(*
	Owns the ended spans of every tracer created from it and hands them to processors.
	Stage the processors every scan, then call tick once; tick passes each ended span to
	every staged processor, releases the span, and clears the staged list.
	The sampler decides which ended spans reach the processors; see onEnd.

	Example:
	provider.stageProcessor(consoleProcessor);
	// ... tracers start and end spans ...
	provider.tick(failureReason => reason);
*)
FUNCTION_BLOCK FB_TracerProvider
VAR
	_resource: REFERENCE TO FB_Resource;  // borrowed; the declaring scope owns its lifetime
	_idGenerator: REFERENCE TO FB_IdGenerator_Base;  // borrowed; the declaring scope owns its lifetime
	_sampler: REFERENCE TO FB_Sampler;  // borrowed; the declaring scope owns its lifetime
	_spans: FB_SpanQueue(TcOtlp_GVL.MAX_SPAN_RECORDS_PER_SCAN);  // ended spans waiting to be processed
	_head: POINTER TO ST_LinkedListNode;  // staged processors; the nodes are owned, the processors borrowed
	_failureReason: E_TracerProviderFailureReason;  // first staging failure since the last tick
END_VAR
VAR_OUTPUT
	stagedProcessorCount: UDINT;
END_VAR

(* Releases the staged-list nodes. The processors themselves are borrowed and untouched. *)
METHOD _freeProcessors
VAR
	_idx: UDINT;
	_node: POINTER TO ST_LinkedListNode;
END_VAR
FOR _idx := 0 TO TcOtlp_GVL.MAX_LOOP_COUNT DO
	IF THIS^._head = 0 THEN
		EXIT;
	END_IF
	_node := THIS^._head^.nxt;
	__DELETE(THIS^._head);
	THIS^._head := _node;
	// count down per node, so the count never claims nodes that are gone or hides ones that remain
	IF THIS^.stagedProcessorCount > 0 THEN
		THIS^.stagedProcessorCount := THIS^.stagedProcessorCount - 1;
	END_IF
END_FOR
END_METHOD

METHOD FB_Exit : BOOL
VAR_INPUT
	bInCopyCode: BOOL;  // TRUE: the exit method is called in order to leave the instance which will be copied afterwards (online change).
END_VAR
IF NOT bInCopyCode THEN
	THIS^._freeProcessors();
END_IF
END_METHOD

//FB_Init is always available implicitly and it is used primarily for initialization.
//The return value is not evaluated. For a specific influence, you can also declare the
//methods explicitly and provide additional code there with the standard initialization
//code. You can evaluate the return value.
METHOD FB_Init: BOOL
VAR_INPUT
    bInitRetains: BOOL; // TRUE: the retain variables are initialized (reset warm / reset cold)
    bInCopyCode: BOOL;  // TRUE: the instance will be copied to the copy code afterward (online change)
	resource: REFERENCE TO FB_Resource;
	idGenerator: REFERENCE TO FB_IdGenerator_Base;  // the source of identifiers for every tracer of this provider
	sampler: REFERENCE TO FB_Sampler;  // decides which spans are sampled; TcOtlp_GVL.defaultSampler is the OpenTelemetry default
END_VAR
THIS^._resource REF= resource;
THIS^._idGenerator REF= idGenerator;
THIS^._sampler REF= sampler;
END_METHOD

(*
	Takes ownership of an ended span and queues it for processing. On success pSpan is
	cleared; on failure it is left unchanged and still owned by the caller.
	A span that is not sampled is released instead, and that counts as success. The sampler's
	onEnd is asked only about spans that are still sampled, so it can drop a span but never
	keep one that its onStart dropped.
*)
METHOD onEnd : BOOL
VAR_IN_OUT
	pSpan: POINTER TO FB_Span;
END_VAR
VAR
	_pushFailureReason: E_SpanQueueFailureReason;
END_VAR
IF pSpan = 0 THEN
	RETURN;
END_IF

IF pSpan^.isSampled() THEN
	THIS^.sampler.onEnd(span:=pSpan^);
END_IF

IF NOT pSpan^.isSampled() THEN
	pSpan^.delete(pSelf:=pSpan);
	onEnd := TRUE;
	RETURN;
END_IF

onEnd := THIS^._spans.push(pValue:=pSpan, failureReason=>_pushFailureReason);
END_METHOD

(*
	Adds a processor for the next tick. The processor is borrowed and must outlive the tick.
	Staging the same processor twice has no effect. At most MAX_LOOP_COUNT processors can be
	staged per tick; staging more fails with STAGE_PROCESSOR_FAILURE. Returns the provider so
	calls can chain.
*)
METHOD stageProcessor : REFERENCE TO FB_TracerProvider
VAR_INPUT
	processor: REFERENCE TO FB_SpanProcessor_Base;
END_VAR
VAR
	_idx: UDINT;
	_node: POINTER TO ST_LinkedListNode;
END_VAR
stageProcessor REF= THIS^;

IF NOT __ISVALIDREF(processor) THEN
	RETURN;
END_IF

IF THIS^._head = 0 THEN
	THIS^._head := __NEW(ST_LinkedListNode);
	IF THIS^._head = 0 THEN
		THIS^._failureReason := E_TracerProviderFailureReason.STAGE_PROCESSOR_FAILURE;
		RETURN;
	END_IF
	THIS^._head^.val := processor.pSelf;
	THIS^.stagedProcessorCount := 1;
	RETURN;
END_IF

_node := THIS^._head;
FOR _idx := 0 TO TcOtlp_GVL.MAX_LOOP_COUNT DO
	IF _node^.val = processor.pSelf THEN
		RETURN;
	ELSIF _node^.nxt = 0 THEN
		// at most MAX_LOOP_COUNT nodes, so _freeProcessors always releases them all
		IF THIS^.stagedProcessorCount >= TcOtlp_GVL.MAX_LOOP_COUNT THEN
			THIS^._failureReason := E_TracerProviderFailureReason.STAGE_PROCESSOR_FAILURE;
			RETURN;
		END_IF
		_node^.nxt := __NEW(ST_LinkedListNode);
		IF _node^.nxt = 0 THEN
			THIS^._failureReason := E_TracerProviderFailureReason.STAGE_PROCESSOR_FAILURE;
			RETURN;
		END_IF
		_node^.nxt^.val := processor.pSelf;
		THIS^.stagedProcessorCount := THIS^.stagedProcessorCount + 1;
		RETURN;
	END_IF
	_node := _node^.nxt;
END_FOR
END_METHOD

(*
	Call once per scan, after staging processors. Passes every queued ended span to each staged
	processor in staging order, releases the span, then ticks the processors and the id
	generator. The queue and the staged list are always cleared, so spans are never carried
	into the next scan: with no processors staged they are released unprocessed.
*)
METHOD tick : BOOL
VAR_OUTPUT
	failureReason: E_TracerProviderFailureReason;
END_VAR
VAR
	_i: UDINT;
	_j: UDINT;
	_count: UDINT;
	_node: POINTER TO ST_LinkedListNode;
	_processor: POINTER TO FB_SpanProcessor_Base;
	_span: POINTER TO FB_Span;
	_popFailureReason: E_SpanQueueFailureReason;
	_idGenFailureReason: E_IdGenFailureReason;
END_VAR
failureReason := THIS^._failureReason;
IF failureReason <> E_TracerProviderFailureReason.NA THEN
	JMP _endLabel;
END_IF

// hand each ended span to every staged processor, then release it
_count := THIS^._spans.count;
FOR _i := 1 TO _count DO
	IF NOT THIS^._spans.pop(pValue:=_span, failureReason=>_popFailureReason) THEN
		failureReason := E_TracerProviderFailureReason.QUEUE_POP_FAILURE;
		JMP _endLabel;
	END_IF
	_node := THIS^._head;
	FOR _j := 1 TO THIS^.stagedProcessorCount DO
		IF _node = 0 THEN
			failureReason := E_TracerProviderFailureReason.UNEXPECTED_NULL_LINKED_LIST_NODE;
			JMP _endLabel;
		END_IF
		_processor := _node^.val;
		IF _processor = 0 THEN
			failureReason := E_TracerProviderFailureReason.UNEXPECTED_NULL_PROCESSOR_POINTER;
			JMP _endLabel;
		END_IF
		_processor^.onEnd(_span^);
		_node := _node^.nxt;
	END_FOR
	_span^.delete(pSelf:=_span);
END_FOR

// tick each processor
_node := THIS^._head;
FOR _j := 1 TO THIS^.stagedProcessorCount DO
	IF _node = 0 THEN
		failureReason := E_TracerProviderFailureReason.UNEXPECTED_NULL_LINKED_LIST_NODE;
		JMP _endLabel;
	END_IF
	_processor := _node^.val;
	IF _processor = 0 THEN
		failureReason := E_TracerProviderFailureReason.UNEXPECTED_NULL_PROCESSOR_POINTER;
		JMP _endLabel;
	END_IF
	_processor^.tick();
	_node := _node^.nxt;
END_FOR

_endLabel:
IF _span <> 0 THEN _span^.delete(pSelf:=_span); END_IF
THIS^._spans.free();
THIS^._freeProcessors();
THIS^._failureReason := E_TracerProviderFailureReason.NA;

// refill the identifier buffer for the next scan
IF __ISVALIDREF(THIS^._idGenerator)
	AND_THEN NOT THIS^._idGenerator.tick(failureReason=>_idGenFailureReason)
	AND_THEN failureReason = E_TracerProviderFailureReason.NA THEN
	failureReason := E_TracerProviderFailureReason.ID_GENERATOR_TICK_FAILURE;
END_IF

tick := failureReason = E_TracerProviderFailureReason.NA;
END_METHOD

PROPERTY idGenerator : REFERENCE TO FB_IdGenerator_Base
GET
idGenerator REF= THIS^._idGenerator;
END_GET
END_PROPERTY

PROPERTY resource : REFERENCE TO FB_Resource
GET
resource REF= THIS^._resource;
END_GET
END_PROPERTY

(* The sampler given to FB_Init, or TcOtlp_GVL.defaultSampler if that reference is invalid. *)
PROPERTY sampler : REFERENCE TO FB_Sampler
GET
IF __ISVALIDREF(THIS^._sampler) THEN
	sampler REF= THIS^._sampler;
ELSE
	sampler REF= TcOtlp_GVL.defaultSampler;
END_IF
END_GET
END_PROPERTY

END_FUNCTION_BLOCK

(* stored: Version 1.1.0.1
   POU FB_TracerProvider: Id {b48a75f0-4a41-4530-9577-d77afb3ee72b}, SpecialFunc None
   Method _freeProcessors: Id {7d098421-3f28-4074-b093-7b198fc76f6e}
   Method FB_Exit: Id {3862a08d-ca0c-4c94-87c9-51375cc5ca7c}
   Method FB_Init: Id {f6a38c97-a50d-4983-a41a-6e702d6849d7}
   Method onEnd: Id {0aaebea3-418a-4f50-b3b0-6f1a94c96d96}
   Method stageProcessor: Id {0ae7d757-2fa4-42cf-bb9a-edd28ebf84dd}
   Method tick: Id {4389ed7d-6a44-4760-adbb-ad0ad20dbd16}
   Property idGenerator: Id {a262f1da-df4d-43ee-84b6-b44c18153b89}
   Get Get: Id {29c6ea03-2912-4ac7-b025-35809fb995cf}
   Property resource: Id {fdb15dde-91d3-4ead-9c92-52fca49b1d49}
   Get Get: Id {bbfec233-bb62-41c1-94c6-632763a36ebc}
   Property sampler: Id {33b6b075-deed-496d-bb0b-7e81c1bfe2e7}
   Get Get: Id {65cd22d8-90df-4796-87be-ce24b5fd71ec} *)
